(* IEC 61131-3 sources: plc-st-coding-agent/progress/f14_agent_v14/release/datasets/selfmade/tests, 15 files *)

(* ---- self-easy-01.reference.st ---- *)
FUNCTION_BLOCK FB
VAR_INPUT
    enable : BOOL;
    values : ARRAY[1..8] OF INT;
    count : INT;
    avgEnable : BOOL;
END_VAR
VAR_OUTPUT
    avgOut : REAL;
END_VAR
VAR
    i : INT;
    n : INT;
    sum : DINT;
    keep : REAL;
END_VAR

(* 先把有效样本数裁剪到 [0, 8]，负数和超长都收敛到合法范围 *)
n := count;
IF n < 0 THEN
    n := 0;
ELSIF n > 8 THEN
    n := 8;
END_IF

(* 要点：输出变量在每周期扫描开头就被赋成本周期的计算结果，
   "保持不变"没法靠"不写它"实现——必须先读回旧值再决定写不写。
   这里用静态变量 keep 记住上一周期的有效结果。 *)
IF enable AND avgEnable AND n > 0 THEN
    sum := 0;
    FOR i := 1 TO n DO
        sum := sum + values[i];
    END_FOR
    keep := DINT_TO_REAL(sum) / INT_TO_REAL(n);
END_IF
avgOut := keep;
END_FUNCTION_BLOCK

(* ---- self-easy-02.reference.st ---- *)
FUNCTION_BLOCK FB
VAR_INPUT
    tankLevel : REAL;
    outletFlow : REAL;
    inletPermit : BOOL;
    resetBtn : BOOL;
END_VAR
VAR_OUTPUT
    pumpRun : BOOL;
    alarmHigh : BOOL;
    alarmLow : BOOL;
    outletValveOpen : BOOL;
END_VAR
VAR
    resetPrev : BOOL;
    resetEdge : BOOL;
    latchReset : BOOL;
END_VAR

(* 复位只取上升沿：按住不放只生效一次。
   边沿必须用独立的 prev 变量记忆上一拍电平，不能写成
   "resetEdge := resetBtn AND NOT resetEdge" —— 那是拿输出当记忆，
   按钮按住时 resetEdge 会振成 真/假/真/假，每两拍就多一个假边沿。 *)
resetEdge := resetBtn AND NOT resetPrev;
resetPrev := resetBtn;
latchReset := resetEdge;

(* 报警自保持：置位优先于复位，且复位条件只在上升沿成立一个周期 *)
(* 置位**不受复位抑制**：报警条件是硬联锁，按下复位不能让它少报一拍。
   复位只在"条件已经消失"时才允许清除（见下面的 gate），两条合起来
   才等价于第 5 条"报警优先于复位"。 *)
IF tankLevel >= 85.0 THEN
    alarmHigh := TRUE;
END_IF
(* 复位只在**条件已经消失**时生效：否则复位当拍会出现
   "液位仍 <= 15 但 alarmLow 已清、出口阀随即打开"的空窗期，
   直接违反"报警优先于复位"这一条。这个洞是模型检查找出来的，
   用例表当时是全绿的。 *)
IF latchReset AND tankLevel < 85.0 THEN
    alarmHigh := FALSE;
END_IF
IF tankLevel <= 15.0 THEN
    alarmLow := TRUE;
END_IF
IF latchReset AND tankLevel > 15.0 THEN
    alarmLow := FALSE;
END_IF

(* 联锁：任一报警存在都不得进料 *)
pumpRun := inletPermit AND NOT alarmHigh AND NOT alarmLow
           AND tankLevel < 85.0 AND tankLevel >= 15.0;

(* 出口阀在低液位报警时强制关闭 *)
outletValveOpen := NOT alarmLow;
END_FUNCTION_BLOCK

(* ---- self-hard-01.reference.st ---- *)
FUNCTION_BLOCK FB
VAR_INPUT
    flowLow : BOOL;
    ackBtn : BOOL;
    sensorOK : BOOL;
END_VAR
VAR_OUTPUT
    alarmActive : BOOL;
    alarmAcked : BOOL;
    highHigh : BOOL;
END_VAR
VAR
    ackPrev : BOOL;
    ackEdge : BOOL;
    acknowledged : BOOL;
END_VAR

ackEdge := ackBtn AND NOT ackPrev;
ackPrev := ackBtn;

(* 高优先级：传感器断线，独立判定，不被低优先级抑制 *)
highHigh := NOT sensorOK;

(* 区分实际确认记忆与输出的“条件消失、待确认清除”标志。 *)
IF flowLow THEN
    IF NOT alarmActive THEN
        acknowledged := FALSE;
    END_IF
    alarmActive := TRUE;
    IF ackEdge THEN
        acknowledged := TRUE;
    END_IF
    alarmAcked := acknowledged;
ELSIF alarmActive THEN
    IF acknowledged OR ackEdge THEN
        alarmActive := FALSE;
        alarmAcked := FALSE;
        acknowledged := FALSE;
    ELSE
        alarmAcked := TRUE;
    END_IF
ELSE
    alarmAcked := FALSE;
    acknowledged := FALSE;
END_IF
END_FUNCTION_BLOCK

(* ---- self-hard-02.reference.st ---- *)
FUNCTION_BLOCK FB
VAR_INPUT
    startBtn : BOOL;
    abortBtn : BOOL;
    setpoint : REAL;
    pv : REAL;
    maxDuration : INT;
END_VAR
VAR_OUTPUT
    elapsed : INT;
    phase : INT;
    timeout : BOOL;
END_VAR
VAR
    startEdgeInputPrev : BOOL;
    startEdge : BOOL;
END_VAR
startEdge := startBtn AND NOT startEdgeInputPrev;
startEdgeInputPrev := startBtn;
IF abortBtn THEN
    phase := 9;
ELSIF startEdge THEN
    phase := 1;
    elapsed := 0;
    timeout := FALSE;
ELSIF phase = 1 OR phase = 2 THEN
    elapsed := elapsed + 1;
    IF elapsed >= maxDuration THEN
        timeout := TRUE;
        phase := 3;
    ELSIF phase = 1 AND pv >= setpoint THEN
        phase := 2;
    END_IF
END_IF
END_FUNCTION_BLOCK

(* ---- self-hard-03.reference.st ---- *)
FUNCTION_BLOCK FB
VAR_INPUT
    pushEn : BOOL;
    pushItem : INT;
    popEn : BOOL;
END_VAR
VAR_IN_OUT
    fifo : ARRAY[1..8] OF INT;
END_VAR
VAR_OUTPUT
    count : INT;
    full : BOOL;
    empty : BOOL;
    head : INT;
END_VAR
VAR
    wasPush : BOOL;
    wasPop : BOOL;
    put : BOOL;
    take : BOOL;
    i : INT;
END_VAR

put := pushEn AND NOT wasPush;
take := popEn AND NOT wasPop;
wasPush := pushEn;
wasPop := popEn;

IF take AND count > 0 THEN
    FOR i := 1 TO count - 1 DO
        fifo[i] := fifo[i + 1];
    END_FOR;
    count := count - 1;
END_IF;
IF put AND count < 8 THEN
    count := count + 1;
    fifo[count] := pushItem;
END_IF;
full := count = 8;
empty := count = 0;
IF empty THEN
    head := 0;
ELSE
    head := fifo[1];
END_IF;
END_FUNCTION_BLOCK

(* ---- self-hard-04.reference.st ---- *)
FUNCTION_BLOCK FB
VAR_INPUT
    demand : INT;
    runHours : ARRAY[1..5] OF LINT;
    rotated : BOOL;
END_VAR
VAR_OUTPUT
    leadPump : INT;
    lagPump : INT;
    runningCount : INT;
END_VAR
VAR
    i : INT;
    need : INT;
    prevNeed : INT;
    best : INT;
    lagMin : INT;
    leadWas : INT;
END_VAR

(* 需求先裁剪到 0..5，否则按泵号取工时可能越界 *)
need := demand;
IF need < 0 THEN
    need := 0;
ELSIF need > 5 THEN
    need := 5;
END_IF
runningCount := need;

(* 全场（工时, 泵号）升序里的第一名：先比工时，工时相同取小泵号 *)
best := 1;
FOR i := 2 TO 5 DO
    IF (runHours[i] < runHours[best]) OR
       ((runHours[i] = runHours[best]) AND (i < best)) THEN
        best := i;
    END_IF
END_FOR

IF need = 0 THEN
    (* 需求归零：主备都清掉，下次正需求重新初选 *)
    leadPump := 0;
    lagPump := 0;
ELSIF leadPump = 0 THEN
    (* 初选：全场最短工时的泵作主泵 *)
    leadPump := best;
ELSE
    (* 迟滞：只有请求有效、且当前主泵比最短工时泵**严格多 50 h 以上**才换主。
       这里刻意不写成"每拍无条件选最短工时"——那样会把迟滞阈值架空，
       每次请求都会立刻换泵，反而加剧磨损与工艺扰动。 *)
    IF rotated AND ((runHours[leadPump] - runHours[best]) > 50) THEN
        leadPump := best;
    END_IF
END_IF

IF need <= 1 THEN
    (* 需求 0/1 台时没有备泵 *)
    lagPump := 0;
ELSE
    (* 备泵：除主泵外的其余泵里（工时, 泵号）最小者 *)
    lagMin := 0;
    FOR i := 1 TO 5 DO
        IF i <> leadPump THEN
            IF lagMin = 0 THEN
                lagMin := i;
            ELSIF (runHours[i] < runHours[lagMin]) OR
                  ((runHours[i] = runHours[lagMin]) AND (i < lagMin)) THEN
                lagMin := i;
            END_IF
        END_IF
    END_FOR
    (* 只在初选、升至需要备泵、或换主时重选备泵，其余拍保留原备泵 *)
    IF (lagPump = 0) OR (lagPump = leadPump) OR (need > prevNeed) OR
       (leadPump <> leadWas) THEN
        lagPump := lagMin;
    END_IF
END_IF

prevNeed := need;
leadWas := leadPump;
END_FUNCTION_BLOCK

(* ---- self-hard-05.reference.st ---- *)
FUNCTION_BLOCK FB
VAR_INPUT
 runRequest : BOOL;
 flameOK : BOOL;
 o2Valid : BOOL;
 o2PV : REAL;
 baseAir : REAL;
 resetBtn : BOOL;
END_VAR
VAR_OUTPUT
 fuelPermit : BOOL;
 trimEnable : BOOL;
 airTrim : REAL;
 airCommand : REAL;
 tripLatched : BOOL;
 o2Fault : BOOL;
END_VAR
VAR
 prevReset : BOOL;
 tripMem : BOOL;
END_VAR
o2Fault := (NOT o2Valid) OR (o2PV < 0.0) OR (o2PV > 21.0);
IF runRequest AND NOT flameOK THEN
 tripMem := TRUE;
ELSIF resetBtn AND NOT prevReset AND NOT runRequest AND NOT flameOK THEN
 tripMem := FALSE;
END_IF;
prevReset := resetBtn;
tripLatched := tripMem;
fuelPermit := runRequest AND flameOK AND NOT tripMem;
trimEnable := fuelPermit AND NOT o2Fault;
IF trimEnable THEN
 airTrim := 2.0 * (2.0 - o2PV);
 IF airTrim > 10.0 THEN airTrim := 10.0; END_IF;
 IF airTrim < -10.0 THEN airTrim := -10.0; END_IF;
ELSE
 airTrim := 0.0;
END_IF;
IF fuelPermit THEN
 airCommand := baseAir + airTrim;
 IF airCommand > 100.0 THEN airCommand := 100.0; END_IF;
 IF airCommand < 0.0 THEN airCommand := 0.0; END_IF;
ELSE
 airCommand := 0.0;
END_IF;
END_FUNCTION_BLOCK

(* ---- self-hard-06.reference.st ---- *)
FUNCTION_BLOCK FB
VAR_INPUT
 runRequest : BOOL;
 pressure : REAL;
 pressureValid : BOOL;
 fuelFlow : REAL;
 steamFlow : REAL;
 outletCmd : INT;
 outletFeedback : INT;
 resetBtn : BOOL;
END_VAR
VAR_OUTPUT
 tripLatched : BOOL;
 fuelPermit : BOOL;
 currentCauseMask : WORD;
 latchedCauseMask : WORD;
 diagnosticActive : BOOL;
END_VAR
VAR
 prevReset : BOOL;
 tripMem : BOOL;
 latMem : WORD;
 valveCnt : INT;
END_VAR
currentCauseMask := 0;
IF resetBtn AND NOT prevReset AND NOT runRequest AND pressureValid
 AND (pressure <= 4200.0) THEN
 tripMem := FALSE;
 latMem := 0;
 valveCnt := 0;
END_IF;
prevReset := resetBtn;
IF NOT runRequest THEN
 valveCnt := 0;
ELSIF NOT pressureValid THEN
 currentCauseMask := 16#0001;
 valveCnt := 0;
 tripMem := TRUE;
ELSIF pressureValid AND (pressure >= 4500.0) THEN
 IF (outletCmd >= 50) AND (outletFeedback <= 10) THEN
  valveCnt := valveCnt + 1;
  IF valveCnt > 3 THEN valveCnt := 3; END_IF;
 ELSE
  valveCnt := 0;
 END_IF;
 IF valveCnt >= 3 THEN
  currentCauseMask := currentCauseMask OR 16#0002;
 END_IF;
 IF (fuelFlow >= 4.0) AND (steamFlow <= 10.0) THEN
  currentCauseMask := currentCauseMask OR 16#0004;
 END_IF;
 IF currentCauseMask = 0 THEN
  currentCauseMask := 16#0008;
 END_IF;
 tripMem := TRUE;
ELSE
 valveCnt := 0;
END_IF;
IF tripMem THEN
 latMem := latMem OR currentCauseMask;
END_IF;
tripLatched := tripMem;
latchedCauseMask := latMem;
diagnosticActive := (currentCauseMask <> 0);
fuelPermit := runRequest AND NOT tripMem;
END_FUNCTION_BLOCK

(* ---- self-hard-07.reference.st ---- *)
FUNCTION_BLOCK FB
VAR_INPUT
 mode : INT;
 resetBtn : BOOL;
 scanSeconds : REAL;
 tempSP : REAL;
 tempPV : REAL;
 flowPV : REAL;
 manualFlowSP : REAL;
 manualValve : REAL;
END_VAR
VAR_OUTPUT
 flowSP : REAL;
 valveCommand : REAL;
 fault : BOOL;
 normalMode : BOOL;
END_VAR
VAR
 prevReset : BOOL;
 initDone : BOOL;
 lastMode : INT;
 accT : REAL;
 accF : REAL;
 oFlow : REAL;
 oValve : REAL;
 eTemp : REAL;
 eFlow : REAL;
 trial : REAL;
 normalMem : BOOL;
END_VAR
fault := (mode < 0) OR (mode > 2) OR (scanSeconds <= 0.0) OR (scanSeconds > 10.0);
normalMem := FALSE;
IF (NOT initDone) OR (resetBtn AND NOT prevReset) OR fault THEN
 oFlow := manualFlowSP;
 oValve := manualValve;
 accT := oFlow - 1.0 * (tempSP - tempPV);
 accF := oValve - 2.0 * (oFlow - flowPV);
 lastMode := mode;
 initDone := TRUE;
ELSIF lastMode <> mode THEN
 IF mode <> 2 THEN
  oFlow := manualFlowSP;
 END_IF;
 accT := oFlow - 1.0 * (tempSP - tempPV);
 accF := oValve - 2.0 * (oFlow - flowPV);
 lastMode := mode;
ELSE
 normalMem := TRUE;
 IF mode = 0 THEN
  oFlow := manualFlowSP;
  oValve := manualValve;
  accT := oFlow - 1.0 * (tempSP - tempPV);
  accF := oValve - 2.0 * (oFlow - flowPV);
 ELSIF mode = 1 THEN
  oFlow := manualFlowSP;
  accT := oFlow - 1.0 * (tempSP - tempPV);
  eFlow := oFlow - flowPV;
  trial := accF + 0.5 * eFlow * scanSeconds;
  oValve := 2.0 * eFlow + trial;
  IF oValve > 100.0 THEN oValve := 100.0; END_IF;
  IF oValve < 0.0 THEN oValve := 0.0; END_IF;
  accF := oValve - 2.0 * eFlow;
 ELSE
  eTemp := tempSP - tempPV;
  trial := accT + 0.2 * eTemp * scanSeconds;
  oFlow := 1.0 * eTemp + trial;
  IF oFlow > 50.0 THEN oFlow := 50.0; END_IF;
  IF oFlow < 0.0 THEN oFlow := 0.0; END_IF;
  accT := oFlow - 1.0 * eTemp;
  eFlow := oFlow - flowPV;
  trial := accF + 0.5 * eFlow * scanSeconds;
  oValve := 2.0 * eFlow + trial;
  IF oValve > 100.0 THEN oValve := 100.0; END_IF;
  IF oValve < 0.0 THEN oValve := 0.0; END_IF;
  accF := oValve - 2.0 * eFlow;
 END_IF;
END_IF;
prevReset := resetBtn;
flowSP := oFlow;
valveCommand := oValve;
normalMode := normalMem;
END_FUNCTION_BLOCK

(* ---- self-medium-01.reference.st ---- *)
(* 配方结构体必须显式定义：题目给的是 ARRAY[1..8] OF ST_Recipe，
   没有 TYPE 块就读不到字段名，结构体成员访问会被直接判错。 *)
TYPE ST_Recipe :
STRUCT
    recipeID : INT;
    totalRatio : REAL;
    temperature : REAL;
END_STRUCT
END_TYPE

FUNCTION_BLOCK FB
VAR_INPUT
    recipe : ARRAY[1..8] OF ST_Recipe;
    selSlot : INT;
    loadCmd : BOOL;
    running : BOOL;
END_VAR
VAR_OUTPUT
    valid : BOOL;
    loadedID : INT;
END_VAR
VAR
    loadPrev : BOOL;
    loadEdge : BOOL;
    ok : BOOL;
    slotOK : BOOL;
    selectedRecipe : ST_Recipe;
END_VAR

loadEdge := loadCmd AND NOT loadPrev;
loadPrev := loadCmd;
(* 生产运行中不接受装载命令：连有效位都不刷新，保持上一次判定 *)
IF loadEdge AND NOT running THEN
    slotOK := (selSlot >= 1) AND (selSlot <= 8);
    (* 关键：先判槽位合法再访问数组。IEC 的 AND 不保证短路，
       所以不能写成 "slotOK AND recipe[selSlot].xxx" 这种依赖短路的写法 *)
    valid := FALSE;
    loadedID := 0;
    IF slotOK THEN
        selectedRecipe := recipe[selSlot];
        ok := selectedRecipe.recipeID <> 0;
        IF selectedRecipe.totalRatio < 99.0 OR selectedRecipe.totalRatio > 101.0 THEN
            ok := FALSE;
        END_IF
        IF selectedRecipe.temperature < 30.0 OR selectedRecipe.temperature > 180.0 THEN
            ok := FALSE;
        END_IF
        valid := ok;
        IF ok THEN
            loadedID := selectedRecipe.recipeID;
        END_IF
    END_IF
END_IF
END_FUNCTION_BLOCK

(* ---- self-medium-02.reference.st ---- *)
FUNCTION_BLOCK FB
VAR_INPUT
    enable : BOOL;
    rawValue : REAL;
END_VAR
VAR_OUTPUT
    filteredValue : REAL;
    windowFull : BOOL;
    sampleCount : INT;
END_VAR
VAR
    buf : ARRAY[1..8] OF REAL;
    wr : INT;
    i : INT;
    sum : REAL;
    keep : REAL;
END_VAR

(* 关断时清空历史，但输出保持最后一次的有效值 *)
IF NOT enable THEN
    FOR i := 1 TO 8 DO
        buf[i] := 0.0;
    END_FOR
    wr := 0;
    sampleCount := 0;
    windowFull := FALSE;
ELSE
    (* 环形缓冲：wr 指向最老元素，写进去就等于淘汰最老的那个 *)
    wr := wr + 1;
    IF wr > 8 THEN
        wr := 1;
    END_IF
    buf[wr] := rawValue;
    IF sampleCount < 8 THEN
        sampleCount := sampleCount + 1;
    END_IF
    windowFull := sampleCount >= 8;

    (* 只对**实际已有**的样本求平均，未满时不得按 0 填充 *)
    sum := 0.0;
    FOR i := 1 TO sampleCount DO
        sum := sum + buf[i];
    END_FOR
    keep := sum / INT_TO_REAL(sampleCount);
END_IF
(* 每一拍都从静态变量刷新输出：输出变量本身不记忆，靠 keep 记忆 *)
filteredValue := keep;
END_FUNCTION_BLOCK

(* ---- self-medium-03.reference.st ---- *)
FUNCTION_BLOCK FB
VAR_INPUT
    openBtn : BOOL;
    closeBtn : BOOL;
    openLimit : BOOL;
    closeLimit : BOOL;
    obstacle : BOOL;
END_VAR
VAR_OUTPUT
    motorUp : BOOL;
    motorDown : BOOL;
    errorFlag : BOOL;
END_VAR
VAR
    state : INT;
    openPrev : BOOL;
    closePrev : BOOL;
    openEdge : BOOL;
    closeEdge : BOOL;
    resetEdge : BOOL;
END_VAR

(* state: 0 idle, 1 opening, 2 closing, 3 latched fault. *)
resetEdge := openBtn AND closeBtn AND NOT (openPrev AND closePrev);
openEdge := openBtn AND NOT openPrev;
closeEdge := closeBtn AND NOT closePrev;
openPrev := openBtn;
closePrev := closeBtn;

IF obstacle THEN
    state := 3;
ELSE
    CASE state OF
        0:
            IF openEdge AND NOT closeBtn AND NOT openLimit THEN
                state := 1;
            ELSIF closeEdge AND NOT openBtn AND NOT closeLimit THEN
                state := 2;
            END_IF;
        1:
            IF openLimit THEN
                state := 0;
            END_IF;
        2:
            IF closeLimit THEN
                state := 0;
            END_IF;
        3:
            IF resetEdge THEN
                state := 0;
            END_IF;
    END_CASE;
END_IF;

motorUp := (state = 1) AND NOT obstacle;
motorDown := (state = 2) AND NOT obstacle;
errorFlag := (state = 3);
END_FUNCTION_BLOCK

(* ---- self-medium-04.reference.st ---- *)
FUNCTION_BLOCK FB
VAR_INPUT
    startBtn : BOOL;
    resetBtn : BOOL;
    doneSensor : BOOL;
    targetVol : REAL;
    flowVol : REAL;
END_VAR
VAR_OUTPUT
    valveOpen : BOOL;
    fillsToday : INT;
END_VAR
VAR
    startPrev : BOOL;
    resetPrev : BOOL;
    startEdge : BOOL;
    resetEdge : BOOL;
    accumulated : REAL;
    filling : BOOL;
    waitAck : BOOL;
END_VAR

startEdge := startBtn AND NOT startPrev;
startPrev := startBtn;
resetEdge := resetBtn AND NOT resetPrev;
resetPrev := resetBtn;

(* 复位最高优先级：清零计数、关阀 *)
IF resetEdge THEN
    fillsToday := 0;
    valveOpen := FALSE;
    filling := FALSE;
    waitAck := FALSE;
    accumulated := 0.0;
ELSE
    (* 运途中重复按启动无效：只在非灌装、非待确认时接受 *)
    (* 待确认期间再按启动：允许直接开灌下一瓶，上一瓶未确认就不计数了 *)
    IF startEdge AND waitAck THEN
        waitAck := FALSE;
    END_IF
    IF startEdge AND NOT filling THEN
        filling := TRUE;
        valveOpen := TRUE;
        accumulated := 0.0;
    END_IF

    IF filling THEN
        accumulated := accumulated + flowVol;
        (* 达到或超过目标立即关阀，用 >= 而不是 > *)
        IF accumulated >= targetVol THEN
            valveOpen := FALSE;
            filling := FALSE;
            waitAck := TRUE;
        END_IF
    END_IF

    (* 计数只在满瓶确认之后发生一次 *)
    IF waitAck AND doneSensor THEN
        IF fillsToday < 32767 THEN
            fillsToday := fillsToday + 1;
        END_IF;
        waitAck := FALSE;
    END_IF
END_IF
END_FUNCTION_BLOCK

(* ---- self-medium-05.reference.st ---- *)
FUNCTION_BLOCK FB
VAR_INPUT
 enable : BOOL;
 resetBtn : BOOL;
 scanSeconds : LREAL;
 steamFlow : LREAL;
 fuelFlow : LREAL;
 steamTemp : LREAL;
 steamPressure : LREAL;
END_VAR
VAR_OUTPUT
 qualified : BOOL;
 dataFault : BOOL;
 qualifiedTon : LREAL;
 fuelTon : LREAL;
 revenue : LREAL;
 cost : LREAL;
 netProfit : LREAL;
END_VAR
VAR
 prevReset : BOOL;
 qTon : LREAL;
 fTon : LREAL;
END_VAR
qualified := (steamTemp >= 447.0) AND (steamTemp <= 453.0)
 AND (steamPressure >= 3750.0) AND (steamPressure <= 3850.0);
dataFault := (scanSeconds <= 0.0) OR (scanSeconds > 10.0)
 OR (steamFlow < 0.0) OR (steamFlow > 90.0)
 OR (fuelFlow < 0.0) OR (fuelFlow > 6.0);
IF resetBtn AND NOT prevReset THEN
 qTon := 0.0;
 fTon := 0.0;
ELSIF enable AND NOT dataFault THEN
 fTon := fTon + fuelFlow * scanSeconds / 1000.0;
 IF qualified THEN
  qTon := qTon + steamFlow * scanSeconds / 1000.0;
 END_IF;
END_IF;
prevReset := resetBtn;
qualifiedTon := qTon;
fuelTon := fTon;
revenue := qTon * 280.0;
cost := fTon * 1500.0;
netProfit := revenue - cost;
END_FUNCTION_BLOCK

(* ---- self-medium-06.reference.st ---- *)
FUNCTION_BLOCK FB
VAR_INPUT
 enable : BOOL;
 resetBtn : BOOL;
 sensorValid : BOOL;
 setpoint : REAL;
 temperature : REAL;
 scanSeconds : REAL;
 bias : REAL;
END_VAR
VAR_OUTPUT
 power : REAL;
 correction : REAL;
 fault : BOOL;
END_VAR
VAR
 prevReset : BOOL;
 prevE : REAL;
 hasHist : BOOL;
 eNow : REAL;
 eDe : REAL;
 xx : REAL;
 yy : REAL;
 mx : REAL;
 zx : REAL;
 px : REAL;
 my : REAL;
 zy : REAL;
 py : REAL;
 wsum : REAL;
 wc : REAL;
 cOut : REAL;
 edgeReset : BOOL;
END_VAR
fault := (NOT sensorValid) OR (scanSeconds <= 0.0) OR (scanSeconds > 10.0);
edgeReset := resetBtn AND NOT prevReset;
IF edgeReset OR (NOT enable) OR fault THEN
 cOut := 0.0;
 hasHist := FALSE;
 prevE := 0.0;
ELSE
 eNow := setpoint - temperature;
 IF hasHist THEN
  eDe := (eNow - prevE) / scanSeconds;
 ELSE
  eDe := 0.0;
 END_IF;
 xx := eNow / 10.0;
 IF xx > 1.0 THEN xx := 1.0; END_IF;
 IF xx < -1.0 THEN xx := -1.0; END_IF;
 yy := eDe / 2.0;
 IF yy > 1.0 THEN yy := 1.0; END_IF;
 IF yy < -1.0 THEN yy := -1.0; END_IF;
 mx := MAX(-xx, 0.0);
 zx := 1.0 - ABS(xx);
 px := MAX(xx, 0.0);
 my := MAX(-yy, 0.0);
 zy := 1.0 - ABS(yy);
 py := MAX(yy, 0.0);
 wsum := mx * my + mx * zy + mx * py + zx * my + zx * zy + zx * py
  + px * my + px * zy + px * py;
 wc := mx * my * (-30.0) + mx * zy * (-20.0) + mx * py * (-10.0)
  + zx * my * (-10.0) + zx * zy * 0.0 + zx * py * 10.0
  + px * my * 10.0 + px * zy * 20.0 + px * py * 30.0;
 IF wsum > 0.0 THEN
  cOut := wc / wsum;
 ELSE
  cOut := 0.0;
 END_IF;
 prevE := eNow;
 hasHist := TRUE;
END_IF;
prevReset := resetBtn;
correction := cOut;
IF edgeReset OR (NOT enable) OR fault THEN
 power := 0.0;
ELSE
 power := bias + cOut;
 IF power > 100.0 THEN power := 100.0; END_IF;
 IF power < 0.0 THEN power := 0.0; END_IF;
END_IF;
END_FUNCTION_BLOCK
